// TIA Portal V19 export
TYPE "Data_Response"
   STRUCT
      "FrequencyOutput (0.01Hz)" : Int;
      "Speed Output (Rpm)" : Int;
      "Current Output (0.01A)" : UInt;
   END_STRUCT;
END_TYPE
